// TIA Portal V19 export
TYPE "PidL.PIDConfig"
   STRUCT
      NegGain : Bool;
      P_Sel : Bool := TRUE;
      I_Sel : Bool := TRUE;
      D_Sel : Bool;
      Gain : Real := 2.0;
      Ti : Real := 20.0;
      Td : Real := 10.0;
      DeadBW : Real;
   END_STRUCT;
END_TYPE
